// TIA Portal V21 export
// export: Created 2026-11-07T15:50:59.8980715Z, ExportSetting WithDefaults, DisplayName Totally Integrated Automation Portal, DisplayVersion V21, DisplayName STEP 7 Professional, DisplayVersion V21, DisplayName STEP 7 Safety, DisplayVersion V21, DisplayName Tech WebApplication, DisplayVersion V21, DisplayName WinCC Basic/Comfort/Advanced, DisplayVersion V21, DisplayName WinCC Unified, DisplayVersion V21
TextList "TL_ListSt"  ListRange=Decimal
  TextListEntry   EntryType=SingleValue, Text="čeka"
  TextListEntry   EntryType=SingleValue, From=1, To=1, Text="gotovo"
  TextListEntry   EntryType=SingleValue, From=2, To=2, Text="preskočeno"
  TextListEntry   EntryType=SingleValue, From=3, To=3, Text="u tijeku"
